(*
    Configuration of FB_AnalogInput16/32. See the block headers.
*)
TYPE ST_AiCfg :
STRUCT
    // Live. Number of values averaged into Status.ValueFiltered, limited to
    // 1..GVL_Param.AI_FILTER_MAX_LENGTH. A change restarts the average.
    FilterSize : DINT := 50;
END_STRUCT
END_TYPE

(* stored: Version 1.1.0.1
   DUT ST_AiCfg: Id {f34c9ac5-780c-4c70-a73f-22a50f864b6c} *)
